(* IEC 61131-3 sources: plc-vscode/tests/st/test-ready/rusty/tests/integration/data/cfc, 13 files *)

(* ---- assigning.st ---- *)
FUNCTION main : DINT
VAR
    x : DINT := 200;
    y : DINT := 100;
    pt : pass_through;
END_VAR
    pt.a := x;
    pt.b := y;
    main := pt.a + pt.b;
END_FUNCTION

(* ---- chained_calls.st ---- *)
FUNCTION main : DINT
VAR
    x : DINT := 2;
    y : DINT := 1;
    adder : myAdder;
END_VAR
    adder.x := x;
    adder.y := y;

    // temp1 := x + y + 1;
    // temp2 := temp1 + y + 1;
    // x := temp1 + temp2 = 2*temp1 + y + 1 = 2x + 2y + 2 + y + 1
    // x := 2x + 3y + 3
    adder();
    main := adder.x;
END_FUNCTION

FUNCTION myAdd : DINT
VAR_INPUT
    a, b : DINT;
END_VAR
    myAdd := a + b;
END_FUNCTION

(* ---- chained_calls_galore.st ---- *)
FUNCTION main : DINT
VAR
    x : DINT := 2;
    y : DINT := 2;
    chainer : ridiculous_chaining;
END_VAR
    chainer(x, y);

    main := chainer.z;
END_FUNCTION

FUNCTION myAdd : DINT
VAR_INPUT
    a, b : DINT;
END_VAR
    myAdd := a + b;
END_FUNCTION

(* ---- conditional_return_block_evaluating_false.st ---- *)
FUNCTION main : DINT
    VAR
        conditional : conditional_return;
    END_VAR

    conditional.a := 0;
    conditional.b := 1;
    conditional.res := 5;
    conditional();

    main := conditional.res;
END_FUNCTION

FUNCTION MyGT : BOOL
    VAR_INPUT
        a, b : DINT;
    END_VAR

    IF a > b THEN
        MyGT := TRUE;
    ELSE
        MyGT := FALSE;
    END_IF
END_FUNCTION

(* ---- conditional_return_block_evaluating_true.st ---- *)
FUNCTION main : DINT
    VAR
        conditional : conditional_return;
    END_VAR

    conditional.a := 1;
    conditional.b := 0;
    conditional.res := 5;
    conditional();

    main := conditional.res;
END_FUNCTION

FUNCTION MyGT : BOOL
    VAR_INPUT
        a, b : DINT;
    END_VAR

    IF a > b THEN
        MyGT := TRUE;
    ELSE
        MyGT := FALSE;
    END_IF
END_FUNCTION

(* ---- conditional_return_evaluating_false.st ---- *)
FUNCTION main : DINT
    VAR
        my_val : DINT := 0;
        conditional : conditional_return;
    END_VAR

    conditional.val := my_val;
    conditional();

    main := conditional.val;
END_FUNCTION

(* ---- conditional_return_evaluating_true.st ---- *)
FUNCTION main : DINT
    VAR
        my_val : DINT := 5;
        conditional : conditional_return;
    END_VAR

    conditional.val := my_val;
    conditional();

    main := conditional.val;
END_FUNCTION

(* ---- conditional_return_evaluating_true_negated.st ---- *)
FUNCTION main : DINT
    VAR
        my_val : DINT := 5;
        conditional : conditional_return;
    END_VAR

    conditional.val := my_val;
    conditional();

    main := conditional.val;
END_FUNCTION

(* ---- connection.st ---- *)
FUNCTION main : DINT
VAR
    value : DINT := 2;
END_VAR
    main := myConnection(value);
;
END_FUNCTION

FUNCTION myAdd : DINT
VAR_INPUT
    a, b : DINT;
END_VAR
    myAdd := a + b;
END_FUNCTION

(* ---- function_returns.st ---- *)
FUNCTION main : DINT
    main := FuncyReturn(111);
END_FUNCTION

(* ---- my_add.st ---- *)
FUNCTION main : DINT
VAR
    x : DINT := 2;
    y : DINT := 1;
    adder : myAdder;
END_VAR
    adder.x := x;
    adder.y := y;

    // x := x + y + 1
    adder();
    main := adder.x;
END_FUNCTION

FUNCTION myAdd : DINT
VAR_INPUT
    a, b : DINT;
END_VAR
    myAdd := a + b;
END_FUNCTION

(* ---- select.st ---- *)
FUNCTION main : DINT
VAR
    x : DINT := 2;
    y : DINT := 1;
    selector : select;
END_VAR
    // x > y ? y : x
    selector(x, y);
    // expecting y
    main := selector.selected;
END_FUNCTION

(* ---- variable_assignment.st ---- *)
FUNCTION main : DINT
VAR
    x : DINT := 10;
    y : DINT := 33333;
    assign : assignment;
END_VAR
    assign.a := x;
    assign.b := y;
    assign();
    // b := a
    main := assign.b;
END_FUNCTION
